FUNCTION FC 1 : VOID
BEGIN
NETWORK
      L 1
      T 100
END_FUNCTION
